(* IEC 61131-3 sources: volt/packages/volt-lsp-iec/test-corpus/awa-palletizer/Device/Plc Logic/Application/Library Manager/L_PLCLoggingAccess, 12 files *)

(* ---- L_TFACILITY.dut ---- *)
TYPE L_TFACILITY :
(
	L_PLC_USER_LOG_SCOPE1 := 512,
	L_PLC_USER_LOG_SCOPE2 := 1024,
	L_PLC_USER_LOG_SCOPE3 := 2048
);
END_TYPE

(* ---- L_TSEVERITY.dut ---- *)
TYPE L_TSEVERITY :
(
	L_LOGFATALERROR := 3,
	L_LOGERROR := 2,
	L_LOGWARNING := 1,
	L_LOGINFORMATION := 0
);
END_TYPE

(* ---- GETBOOLEANPROPERTY.pou ---- *)
FUNCTION GETBOOLEANPROPERTY : BOOL
VAR_INPUT
	STKEY : WSTRING;
END_VAR
END_FUNCTION

(* ---- GETCOMPANY.pou ---- *)
FUNCTION GETCOMPANY : WSTRING
END_FUNCTION

(* ---- GETNUMBERPROPERTY.pou ---- *)
FUNCTION GETNUMBERPROPERTY : DINT
VAR_INPUT
	STKEY : WSTRING;
END_VAR
END_FUNCTION

(* ---- GETTEXTPROPERTY.pou ---- *)
FUNCTION GETTEXTPROPERTY : WSTRING
VAR_INPUT
	STKEY : WSTRING;
END_VAR
END_FUNCTION

(* ---- GETTEXTPROPERTY2.pou ---- *)
FUNCTION GETTEXTPROPERTY2 : POINTER TO WSTRING
VAR_INPUT
	STKEY : WSTRING;
END_VAR
END_FUNCTION

(* ---- GETTITLE.pou ---- *)
FUNCTION GETTITLE : WSTRING
END_FUNCTION

(* ---- GETVERSION.pou ---- *)
FUNCTION GETVERSION : VERSION
END_FUNCTION

(* ---- GETVERSIONPROPERTY.pou ---- *)
FUNCTION GETVERSIONPROPERTY : VERSION
VAR_INPUT
	STKEY : WSTRING;
END_VAR
END_FUNCTION

(* ---- L_ADDLOG.pou ---- *)
FUNCTION L_ADDLOG : BOOL
VAR_INPUT
	ESEVERITY : L_TSeverity;
	EFACILITY : L_TFacility;
	SLOGPAYLOAD : STRING(80);
END_VAR
END_FUNCTION

(* ---- L_ADDLOG2.pou ---- *)
FUNCTION L_ADDLOG2 : BOOL
VAR_INPUT
	ESEVERITY : L_TSeverity;
	UDICOMPONENDID : UDINT;
	SLOGPAYLOAD : STRING(80);
	DWERRORID : DWORD;
	STRLANGUAGETABLE : STRING(80);
END_VAR
END_FUNCTION
